// TIA Portal V21 export
// export: Created 2026-11-11T00:48:23.4796283Z, ExportSetting WithDefaults, DisplayName Totally Integrated Automation Portal, DisplayVersion V21 Update 3, DisplayName STEP 7 Professional, DisplayVersion V21 Update 3, DisplayName STEP 7 Safety, DisplayVersion V21, DisplayName Tech WebApplication, DisplayVersion V21, DisplayName WinCC Basic/Comfort/Advanced, DisplayVersion V21 Update 3, DisplayName WinCC Unified, DisplayVersion V21 Update 3
FUNCTION_BLOCK "FB_Scl_sl113"   // FB197, SCL
{ S7_Optimized_Access := 'TRUE' }
VERSION : 0.1
// stored: AutoNumber true, IsIECCheckEnabled false, IsRetainMemResEnabled false, MemoryReserve 100, SetENOAutomatically false, UDAEnableTagReadback false
   VAR_INPUT
      v_cmd : Bool;
      v_o_fb : Bool;
      v_c_fb : Bool;
   END_VAR
   VAR_OUTPUT
      v_q : Bool;
      v_oa : Bool;
      v_ca : Bool;
   END_VAR
   VAR
      inst { S7_SetPoint := 'True'} : DCAT;
   END_VAR
BEGIN
   #inst(CMD := #v_cmd, O_FB := #v_o_fb, C_FB := #v_c_fb, Q => #v_q, OA => #v_oa, CA => #v_ca);
END_FUNCTION_BLOCK
